SUBAPPLICATION logiBUS_AI_MVA_OPC (* logiBUS_AI_MVA (Analog-Eingang in mV) auf VT-Zahlenfeld + OPC-UA (mV als DWORD, ein Kanal) *)
  (* Standard: 61499-2; Description: Copyright (c) 2026 Meisterschulen am Ostbahnhof This program and the accompanying materials are made available under the terms of the Eclipse Public License 2.0 which is available at https://www.eclipse.org/legal/epl-2.0/ SPDX-License-Identifier: EPL-2.0 *)
  (* Version 1.0, 2026-11-15, Franz Höpfinger, Meisterschulen am Ostbahnhof, initial API and implementation and/or initial documentation *)
  PACKAGE MyLib::sys;
  IMPORT isobus::UT::Q::const::IDs::ID_NULL;
  IMPORT logiBUS::io::AI::logiBUS_AI;
  IMPORT logiBUS::io::AI::logiBUS_AI_S;
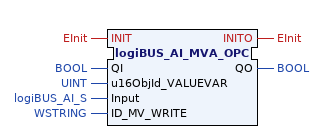
  EVENT_INPUT
    INIT : EInit; (* Initialization Request *)
  END_EVENT
  EVENT_OUTPUT
    INITO : EInit; (* Initialization Confirm *)
  END_EVENT
  VAR_INPUT
    QI : BOOL := TRUE; (* Quality Input - TRUE to enable service *)
    u16ObjId_VALUEVAR : UINT := ID_NULL; (* Object ID CNumberVariable (Spannung in mV) *)
    Input : logiBUS::io::AI::logiBUS_AI_S := logiBUS_AI::Invalid; (* Identify the Input AnalogInput_I1..I8 *)
    ID_MV_WRITE : WSTRING; (* mV-Rueckmelde-Adresse (DWORD, ACTION=PUBLISH) *)
  END_VAR
  VAR_OUTPUT
    QO : BOOL; (* Quality Output - TRUE if service executed successfully *)
  END_VAR
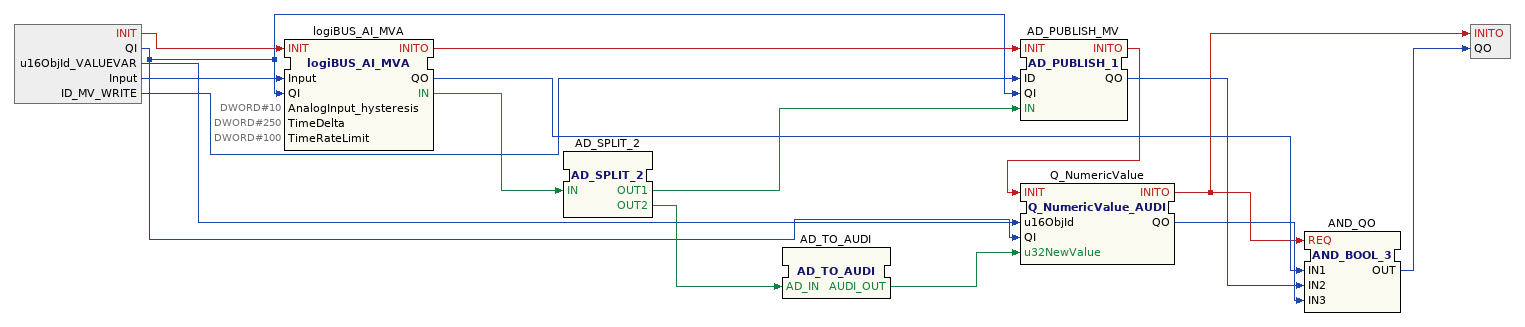
  FBS
    logiBUS_AI_MVA : logiBUS::io::AI::logiBUS_AI_MVA(AnalogInput_hysteresis := DWORD#10, TimeDelta := DWORD#250, TimeRateLimit := DWORD#100);
    AD_SPLIT_2 : adapter::events::unidirectional::AD_SPLIT_2;
    AD_PUBLISH_MV : adapter::net::AD_PUBLISH_1;
    AD_TO_AUDI : adapter::conversion::unidirectional::AD_TO_AUDI;
    Q_NumericValue : isobus::UT::Q::Q_NumericValue_AUDI;
    AND_QO : iec61131::booleanOperators::AND_BOOL_3;
  END_FBS
  EVENT_CONNECTIONS
    INIT TO logiBUS_AI_MVA.INIT;
    logiBUS_AI_MVA.INITO TO AD_PUBLISH_MV.INIT;
    AD_PUBLISH_MV.INITO TO Q_NumericValue.INIT;
    Q_NumericValue.INITO TO INITO;
    Q_NumericValue.INITO TO AND_QO.REQ;
  END_CONNECTIONS
  DATA_CONNECTIONS
    Input TO logiBUS_AI_MVA.Input;
    u16ObjId_VALUEVAR TO Q_NumericValue.u16ObjId;
    ID_MV_WRITE TO AD_PUBLISH_MV.ID;
    QI TO logiBUS_AI_MVA.QI;
    QI TO AD_PUBLISH_MV.QI;
    QI TO Q_NumericValue.QI;
    logiBUS_AI_MVA.QO TO AND_QO.IN1;
    AD_PUBLISH_MV.QO TO AND_QO.IN2;
    Q_NumericValue.QO TO AND_QO.IN3;
    AND_QO.OUT TO QO;
  END_CONNECTIONS
  ADAPTER_CONNECTIONS
    logiBUS_AI_MVA.IN TO AD_SPLIT_2.IN;
    AD_SPLIT_2.OUT1 TO AD_PUBLISH_MV.IN;
    AD_SPLIT_2.OUT2 TO AD_TO_AUDI.AD_IN;
    AD_TO_AUDI.AUDI_OUT TO Q_NumericValue.u32NewValue;
  END_CONNECTIONS
END_SUBAPPLICATION
